DATA_BLOCK "naut_Scan_fast"
{ S7_Optimized_Access := 'TRUE' }
VERSION : 0.1
   VAR
      tags : Struct
         FastDt : LREAL;
      END_STRUCT;
   END_VAR

BEGIN

END_DATA_BLOCK
